(* IEC 61131-3 sources: virtual-bottling-plant/plc/src/machines, 7 files *)

(* ---- FB_Capper.st ---- *)
(* C-501 capper (monoblock with the filler via CV1). Runs a little faster than the filler so
   accumulation conveyors drain after a stop. *)
FUNCTION_BLOCK FB_Capper
  VAR_INPUT
    LineCmd : ST_MachineCmd;
    OwnCmd : E_Command;
    StopReasonCmd : INT;
    HoldId : INT;
    LineHoldId : INT;
    Running : BOOL;
    InputFill : REAL;          (* CV1_Fill, bottles *)
    UpstreamExecute : BOOL;    (* the machine feeding CV1 is producing *)
    OutputFull : BOOL;         (* CV2_Full *)
    Recipe : ST_Recipe;
    NowMs : UDINT;
  END_VAR
  VAR_OUTPUT
    Status : ST_PackagingStatus;
    Run : BOOL;
    SpeedSP : REAL;
  END_VAR
  VAR
    Unit : FB_PackagingUnit;
  END_VAR

  Unit(LineCmd := LineCmd, OwnCmd := OwnCmd, StopReasonCmd := StopReasonCmd, HoldId := HoldId,
       LineHoldId := LineHoldId, Blocked := OutputFull,
       Starved := InputFill < 1.0 AND NOT UpstreamExecute,
       StarvedDelayMs := 2000, Running := Running, NowMs := NowMs);
  Status := Unit.Status;
  Run := Unit.RunOut;
  SpeedSP := Recipe.LineSpeed + 10.0;
END_FUNCTION_BLOCK

(* ---- FB_CasePacker.st ---- *)
(* K-801 case packer, end of line (never blocked). It waits for 6 bottles per case. *)
FUNCTION_BLOCK FB_CasePacker
  VAR_INPUT
    LineCmd : ST_MachineCmd;
    OwnCmd : E_Command;
    StopReasonCmd : INT;
    HoldId : INT;
    LineHoldId : INT;
    Running : BOOL;
    InputFill : REAL;          (* CV4_Fill, bottles *)
    UpstreamExecute : BOOL;    (* the machine feeding CV4 is producing *)
    Recipe : ST_Recipe;
    NowMs : UDINT;
  END_VAR
  VAR_OUTPUT
    Status : ST_PackagingStatus;
    Run : BOOL;
    SpeedSP : REAL;
  END_VAR
  VAR
    Unit : FB_PackagingUnit;
  END_VAR

  Unit(LineCmd := LineCmd, OwnCmd := OwnCmd, StopReasonCmd := StopReasonCmd, HoldId := HoldId,
       LineHoldId := LineHoldId, Blocked := FALSE,
       Starved := InputFill < 6.0 AND NOT UpstreamExecute,
       StarvedDelayMs := 2000, Running := Running, NowMs := NowMs);
  Status := Unit.Status;
  Run := Unit.RunOut;
  SpeedSP := Recipe.LineSpeed / 6.0 + 2.0;  (* cases/min, a little faster than the filler *)
END_FUNCTION_BLOCK

(* ---- FB_Checkweigher.st ---- *)
(* Q-701 checkweigher. Rejects bottles below the fill target minus 10 g (995 g at 1005 g). *)
FUNCTION_BLOCK FB_Checkweigher
  VAR_INPUT
    LineCmd : ST_MachineCmd;
    OwnCmd : E_Command;
    StopReasonCmd : INT;
    HoldId : INT;
    LineHoldId : INT;
    Running : BOOL;
    InputFill : REAL;          (* CV3_Fill, bottles *)
    UpstreamExecute : BOOL;    (* the machine feeding CV3 is producing *)
    OutputFull : BOOL;         (* CV4_Full *)
    Count : UDINT;             (* bottles weighed *)
    RejectCount : UDINT;
    Recipe : ST_Recipe;
    NowMs : UDINT;
  END_VAR
  VAR_OUTPUT
    Status : ST_PackagingStatus;
    Run : BOOL;
    SpeedSP : REAL;
    RejectLimitG : REAL;
    GoodCount : UDINT;
  END_VAR
  VAR
    Unit : FB_PackagingUnit;
  END_VAR

  Unit(LineCmd := LineCmd, OwnCmd := OwnCmd, StopReasonCmd := StopReasonCmd, HoldId := HoldId,
       LineHoldId := LineHoldId, Blocked := OutputFull,
       Starved := InputFill < 1.0 AND NOT UpstreamExecute,
       StarvedDelayMs := 2000, Running := Running, NowMs := NowMs);
  Status := Unit.Status;
  Run := Unit.RunOut;
  SpeedSP := Recipe.LineSpeed + 20.0;
  RejectLimitG := Recipe.FillTargetG - 10.0;
  IF Count >= RejectCount THEN
    GoodCount := Count - RejectCount;
  ELSE
    GoodCount := 0;  (* one counter wrapped before the other *)
  END_IF;
END_FUNCTION_BLOCK

(* ---- FB_Filler.st ---- *)
(* F-401 rotary filler, the line constraint. Interlock PLC-11: it fills only while T-301
   is above its start level (FB_Tank hysteresis), otherwise it is Suspended (starved) with the
   motor off, so it cannot run the buffer dry. *)
FUNCTION_BLOCK FB_Filler
  VAR_INPUT
    LineCmd : ST_MachineCmd;
    OwnCmd : E_Command;
    StopReasonCmd : INT;
    HoldId : INT;
    LineHoldId : INT;
    Running : BOOL;
    OutputFull : BOOL;         (* CV1_Full *)
    BufferPermissive : BOOL;   (* T-301 above the filler start level *)
    Recipe : ST_Recipe;
    NowMs : UDINT;
  END_VAR
  VAR_OUTPUT
    Status : ST_PackagingStatus;
    Run : BOOL;
    SpeedSP : REAL;
    FillTargetG : REAL;
  END_VAR
  VAR
    Unit : FB_PackagingUnit;
  END_VAR

  Unit(LineCmd := LineCmd, OwnCmd := OwnCmd, StopReasonCmd := StopReasonCmd, HoldId := HoldId,
       LineHoldId := LineHoldId, Blocked := OutputFull, Starved := NOT BufferPermissive,
       StarvedDelayMs := 2000, Running := Running, NowMs := NowMs);
  Status := Unit.Status;
  Run := Unit.RunOut AND BufferPermissive;
  SpeedSP := Recipe.LineSpeed;
  FillTargetG := Recipe.FillTargetG;
END_FUNCTION_BLOCK

(* ---- FB_Labeler.st ---- *)
(* L-601 labeler. *)
FUNCTION_BLOCK FB_Labeler
  VAR_INPUT
    LineCmd : ST_MachineCmd;
    OwnCmd : E_Command;
    StopReasonCmd : INT;
    HoldId : INT;
    LineHoldId : INT;
    Running : BOOL;
    InputFill : REAL;          (* CV2_Fill, bottles *)
    UpstreamExecute : BOOL;    (* the machine feeding CV2 is producing *)
    OutputFull : BOOL;         (* CV3_Full *)
    Recipe : ST_Recipe;
    NowMs : UDINT;
  END_VAR
  VAR_OUTPUT
    Status : ST_PackagingStatus;
    Run : BOOL;
    SpeedSP : REAL;
  END_VAR
  VAR
    Unit : FB_PackagingUnit;
  END_VAR

  Unit(LineCmd := LineCmd, OwnCmd := OwnCmd, StopReasonCmd := StopReasonCmd, HoldId := HoldId,
       LineHoldId := LineHoldId, Blocked := OutputFull,
       Starved := InputFill < 1.0 AND NOT UpstreamExecute,
       StarvedDelayMs := 2000, Running := Running, NowMs := NowMs);
  Status := Unit.Status;
  Run := Unit.RunOut;
  SpeedSP := Recipe.LineSpeed + 10.0;
END_FUNCTION_BLOCK

(* ---- FB_LineSequencer.st ---- *)
(* Line start/stop from the local panel (sim operator) or the HMI line command.
   Start: each machine is reset if Stopped, then started once the machine after it is running,
   so the line starts from the case packer back to the filler. Stop: every machine stops.
   Reset: unholds machines whose cause is gone (and resets stopped ones). *)
FUNCTION_BLOCK FB_LineSequencer
  VAR_INPUT
    PbStart : BOOL;
    PbStop : BOOL;
    PbReset : BOOL;
    LineCmd : E_Command;
    F401State : E_PackMLState;
    C501State : E_PackMLState;
    L601State : E_PackMLState;
    Q701State : E_PackMLState;
    K801State : E_PackMLState;
  END_VAR
  VAR_OUTPUT
    F401 : ST_MachineCmd;
    C501 : ST_MachineCmd;
    L601 : ST_MachineCmd;
    Q701 : ST_MachineCmd;
    K801 : ST_MachineCmd;
    StartRequested : BOOL;
  END_VAR
  VAR
    StartEdge : R_TRIG;
    StopEdge : R_TRIG;
    ResetEdge : R_TRIG;
    Stop : BOOL;
    Reset : BOOL;
    Abort : BOOL;
    Clear : BOOL;
  END_VAR

  StartEdge(CLK := PbStart);
  StopEdge(CLK := PbStop);
  ResetEdge(CLK := PbReset);
  Stop := StopEdge.Q OR LineCmd = CMD_STOP;
  Reset := ResetEdge.Q OR LineCmd = CMD_RESET;
  Abort := LineCmd = CMD_ABORT;
  Clear := LineCmd = CMD_CLEAR;

  IF Stop OR Abort THEN
    StartRequested := FALSE;
  ELSIF StartEdge.Q OR LineCmd = CMD_START THEN
    StartRequested := TRUE;
  END_IF;

  K801.Start := StartRequested AND K801State = PML_IDLE;
  Q701.Start := StartRequested AND Q701State = PML_IDLE AND PackMLHasStarted(K801State);
  L601.Start := StartRequested AND L601State = PML_IDLE AND PackMLHasStarted(Q701State);
  C501.Start := StartRequested AND C501State = PML_IDLE AND PackMLHasStarted(L601State);
  F401.Start := StartRequested AND F401State = PML_IDLE AND PackMLHasStarted(C501State);

  K801.Reset := Reset OR (StartRequested AND K801State = PML_STOPPED);
  Q701.Reset := Reset OR (StartRequested AND Q701State = PML_STOPPED);
  L601.Reset := Reset OR (StartRequested AND L601State = PML_STOPPED);
  C501.Reset := Reset OR (StartRequested AND C501State = PML_STOPPED);
  F401.Reset := Reset OR (StartRequested AND F401State = PML_STOPPED);

  K801.Stop := Stop;
  K801.Abort := Abort;
  K801.Clear := Clear;
  Q701.Stop := Stop;
  Q701.Abort := Abort;
  Q701.Clear := Clear;
  L601.Stop := Stop;
  L601.Abort := Abort;
  L601.Clear := Clear;
  C501.Stop := Stop;
  C501.Abort := Abort;
  C501.Clear := Clear;
  F401.Stop := Stop;
  F401.Abort := Abort;
  F401.Clear := Clear;

  (* The request ends once every machine is under way; later stops are not undone. *)
  IF StartRequested AND PackMLHasStarted(F401State) AND PackMLHasStarted(C501State)
     AND PackMLHasStarted(L601State) AND PackMLHasStarted(Q701State)
     AND PackMLHasStarted(K801State) THEN
    StartRequested := FALSE;
  END_IF;
END_FUNCTION_BLOCK

(* ---- FB_LineStatus.st ---- *)
(* Line-level status block: the line is in the state of its constraint machine, F-401. *)
FUNCTION_BLOCK FB_LineStatus
  VAR_INPUT
    FillerState : E_PackMLState;
    Recipe : ST_Recipe;
  END_VAR
  VAR_OUTPUT
    Status : ST_LINEStatus;
  END_VAR

  Status.State := FillerState;
  Status.RecipeId := Recipe.RecipeId;
  Status.RecipeVersion := Recipe.RecipeVersion;
  Status.ProductCode := Recipe.ProductCode;
  (* Lets the bridge see that the PLC program is scanning *)
  Status.PlcHeartbeat := (Status.PlcHeartbeat + 1) MOD 30000;
END_FUNCTION_BLOCK
